Staubli VAL3: _productCycle.pgx

public program _productCycle()
  local bool l_bErr
  local bool l_bStartClock
  local num l_nClock
  local num l_nLastAct
  local num l_nLibIndex
  local string l_sPath
  local bool l_bFound
  local string l_sSelTraj
begin
  while true

    //
    //等待执行命令
    wait(plc:dInExcutePainting==true)
    //获取程序号
    call io:getAnaIO(io:aInItem[0].aAio,rs:nProgCode,l_bErr)
    //搜索对应traj
    call search_traj(l_bFound,l_sSelTraj,rs:nProgCode)
    //如果找到对应的traj，执行traj
    if l_bFound
      call trajectory:makeTraj(l_sSelTraj)
      waitEndMove()
    else
      popUpMsg("未找到喷涂号对应执行程序")
      rs:bIsError=true
      rs:bToStopCycle=true
    endIf
    delay(0)
  endWhile

  //  if l_bStartClock and l_nLastAct!=rs:nActCode
  //    rs:_nCTIndex=(rs:_nCTIndex+1)%size(rs:_nCycleTime)
  //    rs:_nCycleTime[rs:_nCTIndex]=clock()-l_nClock
  //  else
  //    l_bStartClock=true
  //  endIf
  //  l_nClock=clock()
  //  l_nLastAct=rs:nActCode
  //  //delay(0)
  //  //
  //  rs:_nOmacStat=1
  //  rs:sTrajStatus=""
  rs:_sRobotStatus="当前件生产结束"
  //2025.1.6 add 结束扭矩记录程序
  if taskStatus("getForce")!=-1
    delay(0.2)
    taskKill("getForce")
  endIf
end
